SUBAPPLICATION ASRT_AX_SERVER_0_PUBLISH_1 (* Wie adapter::net::ASRT_AX_SERVER_0_CLIENT_1_0, aber lokales PUBLISH_1 statt Remote-CLIENT_1_0 (ein Geraet) *)
  (* Standard: 61499-2; Description: Copyright (c) 2026 HR Agrartechnik GmbH This program and the accompanying materials are made available under the terms of the Eclipse Public License 2.0 which is available at https://www.eclipse.org/legal/epl-2.0/ SPDX-License-Identifier: EPL-2.0 *)
  (* Version 1.2, 2026-11-25, Franz Höpfinger, Meisterschulen am Ostbahnhof, SERVER_0 -> MyLib::net::SERVER_0_QO (IND nur bei QO=TRUE, RSP intern). Ein gescheitertes RSP meldet IND mit QO=FALSE, direkt IND->RSP ergab eine Endlosschleife. *)
  (* Version 1.1, 2026-10-18, Franz Höpfinger, Meisterschulen am Ostbahnhof, Kopie von ASRT_AX_SERVER_0_CLIENT_1_0, CLIENT_1_0 durch PUBLISH_1 ersetzt - als SubAppType, damit FORTE den Typ nicht kennen muss (kein ELF fuer MyLib_AX). SERVER_0: IND direkt auf RSP (sonst bis 4 s Server-Lock fuer alle Publishes) *)
  (* Version 1.0, 2026-09-03, Franz Höpfinger, HR Agrartechnik GmbH, initial API and implementation and/or initial documentation *)
  PACKAGE MyLib::net;
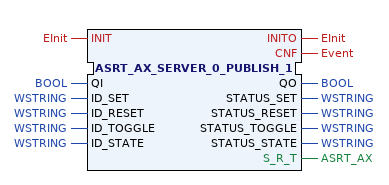
  EVENT_INPUT
    INIT : EInit; (* Initialization *)
  END_EVENT
  EVENT_OUTPUT
    INITO : EInit; (* Initialization Confirm *)
    CNF; (* QO/STATUS updated *)
  END_EVENT
  VAR_INPUT
    QI : BOOL;
    ID_SET : WSTRING; (* Lokale Methodenadresse (ACTION=CREATE_METHOD) fuer den Set-Methodenaufruf *)
    ID_RESET : WSTRING; (* Lokale Methodenadresse (ACTION=CREATE_METHOD) fuer den Reset-Methodenaufruf *)
    ID_TOGGLE : WSTRING; (* Lokale Methodenadresse (ACTION=CREATE_METHOD) fuer den Toggle-Methodenaufruf *)
    ID_STATE : WSTRING; (* Lokale Adresse (ACTION=WRITE) fuer den Zustand *)
  END_VAR
  VAR_OUTPUT
    QO : BOOL; (* TRUE nur wenn SET_SERVER, RESET_SERVER, TOGGLE_SERVER und STATE_CLIENT aktuell alle QO=TRUE melden *)
    STATUS_SET : WSTRING; (* STATUS von SET_SERVER *)
    STATUS_RESET : WSTRING; (* STATUS von RESET_SERVER *)
    STATUS_TOGGLE : WSTRING; (* STATUS von TOGGLE_SERVER *)
    STATUS_STATE : WSTRING; (* STATUS von STATE_CLIENT *)
  END_VAR
  PLUGS
    S_R_T : adapter::types::bidirectional::ASRT_AX; (* Set/Reset/Toggle (in), Zustand (out) *)
  END_PLUGS
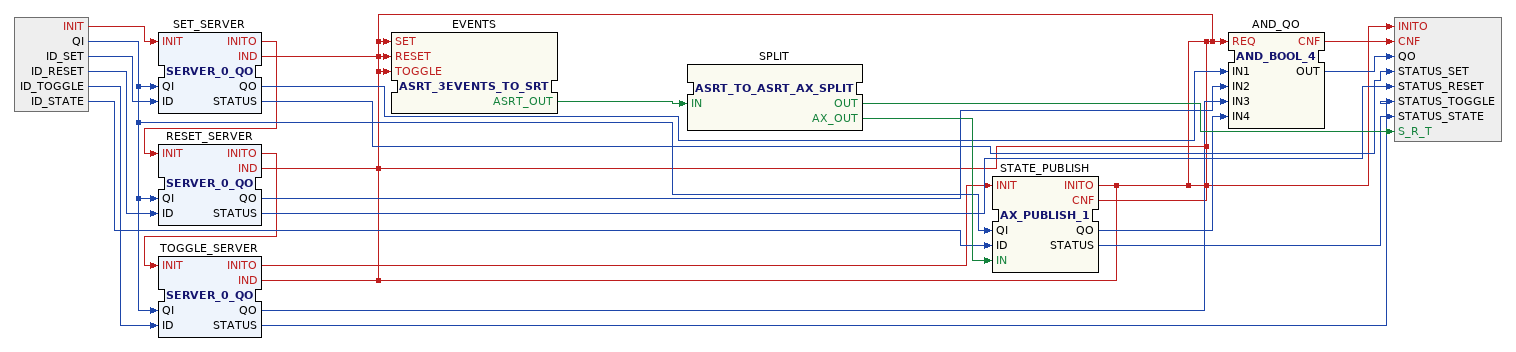
  FBS
    EVENTS : adapter::conversion::unidirectional::ASRT_3EVENTS_TO_SRT;
    SPLIT : adapter::events::bidirectional::ASRT_TO_ASRT_AX_SPLIT;
    STATE_PUBLISH : adapter::net::AX_PUBLISH_1;
    AND_QO : iec61131::booleanOperators::AND_BOOL_4;
  END_FBS
  SUBAPPS
    SET_SERVER : MyLib::net::SERVER_0_QO;
    RESET_SERVER : MyLib::net::SERVER_0_QO;
    TOGGLE_SERVER : MyLib::net::SERVER_0_QO;
  END_SUBAPPS
  EVENT_CONNECTIONS
    INIT TO SET_SERVER.INIT;
    SET_SERVER.INITO TO RESET_SERVER.INIT;
    RESET_SERVER.INITO TO TOGGLE_SERVER.INIT;
    TOGGLE_SERVER.INITO TO STATE_PUBLISH.INIT;
    STATE_PUBLISH.INITO TO INITO;
    STATE_PUBLISH.INITO TO AND_QO.REQ;
    SET_SERVER.IND TO EVENTS.SET;
    SET_SERVER.IND TO AND_QO.REQ;
    RESET_SERVER.IND TO EVENTS.RESET;
    RESET_SERVER.IND TO AND_QO.REQ;
    TOGGLE_SERVER.IND TO EVENTS.TOGGLE;
    TOGGLE_SERVER.IND TO AND_QO.REQ;
    STATE_PUBLISH.CNF TO AND_QO.REQ;
    AND_QO.CNF TO CNF;
  END_CONNECTIONS
  DATA_CONNECTIONS
    QI TO SET_SERVER.QI;
    ID_SET TO SET_SERVER.ID;
    SET_SERVER.QO TO AND_QO.IN1;
    SET_SERVER.STATUS TO STATUS_SET;
    QI TO RESET_SERVER.QI;
    ID_RESET TO RESET_SERVER.ID;
    RESET_SERVER.QO TO AND_QO.IN2;
    RESET_SERVER.STATUS TO STATUS_RESET;
    QI TO TOGGLE_SERVER.QI;
    ID_TOGGLE TO TOGGLE_SERVER.ID;
    TOGGLE_SERVER.QO TO AND_QO.IN3;
    TOGGLE_SERVER.STATUS TO STATUS_TOGGLE;
    QI TO STATE_PUBLISH.QI;
    ID_STATE TO STATE_PUBLISH.ID;
    STATE_PUBLISH.QO TO AND_QO.IN4;
    AND_QO.OUT TO QO;
    STATE_PUBLISH.STATUS TO STATUS_STATE;
  END_CONNECTIONS
  ADAPTER_CONNECTIONS
    EVENTS.ASRT_OUT TO SPLIT.IN;
    SPLIT.OUT TO S_R_T;
    SPLIT.AX_OUT TO STATE_PUBLISH.IN;
  END_CONNECTIONS
END_SUBAPPLICATION
